Staubli VAL3: createUserTask.pgx

program createUserTask()
begin
  //作用：调用自定义的任务
  //1.创建动作Action任务
  call act:create()
  //2.创建视觉任务
end
